FUNCTION_BLOCK SingleSolenoidCylinder EXTENDS ActuatorBase
VAR
    _Solenoid        : REFERENCE TO BOOL;
    _ExtendedSensor  : REFERENCE TO BOOL;
    _RetractedSensor : REFERENCE TO BOOL;
END_VAR
(*
    SingleSolenoidCylinder

    One solenoid with spring return: energized extends, de-energized retracts.
    An end sensor at each end.
*)

METHOD FB_init : BOOL
VAR_INPUT
    bInitRetains    : BOOL;
    bInCopyCode     : BOOL;
    Name            : STRING(32);
    MoveTimeout     : TIME;
    Solenoid        : REFERENCE TO BOOL;
    ExtendedSensor  : REFERENCE TO BOOL;
    RetractedSensor : REFERENCE TO BOOL;
END_VAR
_Solenoid REF= Solenoid;
_ExtendedSensor REF= ExtendedSensor;
_RetractedSensor REF= RetractedSensor;
Configure(Name := Name, MoveTimeout := MoveTimeout);
END_METHOD

METHOD PROTECTED IsWired : BOOL
IsWired := __ISVALIDREF(_Solenoid) AND __ISVALIDREF(_ExtendedSensor) AND __ISVALIDREF(_RetractedSensor);
END_METHOD

METHOD PROTECTED DriveOutputs
VAR_INPUT
    Target : E_ActuatorTarget;
END_VAR
_Solenoid := Target = E_ActuatorTarget.Extended;   // anything else: the spring retracts it
END_METHOD

METHOD PROTECTED IsAtPosition : BOOL
VAR_INPUT
    Position : E_ActuatorTarget;
END_VAR
CASE Position OF
    E_ActuatorTarget.Extended:
        IsAtPosition := _ExtendedSensor AND NOT _RetractedSensor;
    E_ActuatorTarget.Retracted:
        IsAtPosition := _RetractedSensor AND NOT _ExtendedSensor;
ELSE
    IsAtPosition := FALSE;
END_CASE
END_METHOD

METHOD PROTECTED DriveSafe
_Solenoid := FALSE;                                 // the spring takes it to the retracted end
END_METHOD

END_FUNCTION_BLOCK

(* stored: Version 1.1.0.1, ProductVersion 3.1.4026.0
   POU SingleSolenoidCylinder: Id {9610f7f6-417e-49aa-a504-132e889d69c2}, SpecialFunc None
   Method FB_init: Id {8cf15dde-2733-4f49-b7d8-4ca428e47aef}
   Method IsWired: Id {4849c915-07d7-42fc-9d03-fde1775a6d48}
   Method DriveOutputs: Id {e070fba6-06e9-4fe5-b145-92f150b1f980}
   Method IsAtPosition: Id {6488f2df-2cb5-439c-a2af-aa5aee8e373b}
   Method DriveSafe: Id {dc00bd41-8f51-4fd3-929b-f2373061473e} *)
